(* IEC 61131-3 sources: plcassist-cli/packages/volt-lsp-iec/test-corpus/bakon-nano/Device/Plc Logic/Application/Library Manager/CmpBinTagUtilIec, 34 files *)

(* ---- BTAGALIGNMENTS.gvl ---- *)
VAR_GLOBAL
	ALIGN42 : BTagAlignment := STRUCT(uiModulus := 4, uiRemainder := 2);
	ALIGN40 : BTagAlignment := STRUCT(uiModulus := 4, uiRemainder := 0);
END_VAR

(* ---- RETURNVALUES.gvl ---- *)
VAR_GLOBAL
	ERR_OK : UDINT := 16#0;
	ERR_FAILED : UDINT := 16#1;
	ERR_PARAMETER : UDINT := 16#2;
	ERR_NOTIMPLEMENTED : UDINT := 16#C;
	ERR_NOMEMORY : UDINT := 16#11;
	ERR_BTAG_TAGOVERLAP : UDINT := 16#400;
	ERR_BTAG_BUFFEROVERRUN : UDINT := 16#401;
	ERR_BTAG_MAXNESTINGDEPTH : UDINT := 16#402;
	ERR_BTAG_NOTAG : UDINT := 16#403;
	ERR_BTAG_NODATATAG : UDINT := 16#404;
	ERR_BTAG_NOCONTAINERTAG : UDINT := 16#405;
	ERR_BTAG_NOTTOPLEVEL : UDINT := 16#406;
	ERR_BTAG_ALIGNMENT : UDINT := 16#407;
	INVALID_HANDLE : __UXINT := RTS_INVALID_HANDLE;
END_VAR

(* ---- BTAGREADERCREATE.fun ---- *)
FUNCTION BTAGREADERCREATE : RTS_IEC_HANDLE
VAR_INPUT
	PBUFFER : POINTER TO BYTE;
	DWSIZE : DWORD;
	PRESULT : POINTER TO RTS_IEC_RESULT;
END_VAR
END_FUNCTION

(* ---- BTAGREADERCREATEDYNAMIC.fun ---- *)
FUNCTION BTAGREADERCREATEDYNAMIC : RTS_IEC_HANDLE
VAR_INPUT
	PRESULT : POINTER TO RTS_IEC_RESULT;
END_VAR
END_FUNCTION

(* ---- BTAGREADERDESTROY.fun ---- *)
FUNCTION BTAGREADERDESTROY : RTS_IEC_RESULT
VAR_INPUT
	HREADER : RTS_IEC_HANDLE;
END_VAR
END_FUNCTION

(* ---- BTAGREADERGETCOMPLEXCONTENT.fun ---- *)
FUNCTION BTAGREADERGETCOMPLEXCONTENT : RTS_IEC_RESULT
VAR_INPUT
	HREADER : RTS_IEC_HANDLE;
	PPBUFFER : POINTER TO POINTER TO BYTE;
	PULSIZE : POINTER TO UDINT;
END_VAR
END_FUNCTION

(* ---- BTAGREADERGETCONTENT.fun ---- *)
FUNCTION BTAGREADERGETCONTENT : RTS_IEC_RESULT
VAR_INPUT
	HREADER : RTS_IEC_HANDLE;
	PPBUFFER : POINTER TO POINTER TO BYTE;
	PULSIZE : POINTER TO UDINT;
END_VAR
END_FUNCTION

(* ---- BTAGREADERGETSTRING.fun ---- *)
FUNCTION BTAGREADERGETSTRING : RTS_IEC_RESULT
VAR_INPUT
	HREADER : RTS_IEC_HANDLE;
	PPBUFFER : POINTER TO POINTER TO BYTE;
	PULSIZE : POINTER TO UDINT;
	BADDENDOFSTRING : BOOL;
END_VAR
END_FUNCTION

(* ---- BTAGREADERGETTAGID.fun ---- *)
FUNCTION BTAGREADERGETTAGID : RTS_IEC_RESULT
VAR_INPUT
	HREADER : RTS_IEC_HANDLE;
	PULTAGID : POINTER TO UDINT;
END_VAR
END_FUNCTION

(* ---- BTAGREADERGETTAGLEN.fun ---- *)
FUNCTION BTAGREADERGETTAGLEN : RTS_IEC_RESULT
VAR_INPUT
	HREADER : RTS_IEC_HANDLE;
	PULTAGLEN : POINTER TO UDINT;
END_VAR
END_FUNCTION

(* ---- BTAGREADERINIT.fun ---- *)
FUNCTION BTAGREADERINIT : RTS_IEC_RESULT
VAR_INPUT
	HREADER : RTS_IEC_HANDLE;
	PBUFFER : POINTER TO BYTE;
	DWBUFFERSIZE : DWORD;
END_VAR
END_FUNCTION

(* ---- BTAGREADERISDATATAG.fun ---- *)
FUNCTION BTAGREADERISDATATAG : RTS_IEC_RESULT
VAR_INPUT
	HREADER : RTS_IEC_HANDLE;
	PBDATATAG : POINTER TO BOOL;
END_VAR
END_FUNCTION

(* ---- BTAGREADERMOVENEXT.fun ---- *)
FUNCTION BTAGREADERMOVENEXT : RTS_IEC_RESULT
VAR_INPUT
	HREADER : RTS_IEC_HANDLE;
	PNELEMENTTYPE : POINTER TO BTagElementType;
END_VAR
END_FUNCTION

(* ---- BTAGREADERPEEKNEXT.fun ---- *)
FUNCTION BTAGREADERPEEKNEXT : BTagElementType
VAR_INPUT
	HREADER : RTS_IEC_HANDLE;
END_VAR
END_FUNCTION

(* ---- BTAGREADERSKIPCONTENT.fun ---- *)
FUNCTION BTAGREADERSKIPCONTENT : RTS_IEC_RESULT
VAR_INPUT
	HREADER : RTS_IEC_HANDLE;
END_VAR
END_FUNCTION

(* ---- BTAGSWAPHEADER.fun ---- *)
FUNCTION BTAGSWAPHEADER : DWORD
VAR_INPUT
	PHEADERTAG : POINTER TO DWORD;
	BSWAP : DINT;
END_VAR
END_FUNCTION

(* ---- BTAGWRITERAPPENDBLOB.fun ---- *)
FUNCTION BTAGWRITERAPPENDBLOB : RTS_IEC_RESULT
VAR_INPUT
	HWRITER : RTS_IEC_HANDLE;
	PDATA : POINTER TO BYTE;
	DWDATASIZE : DWORD;
END_VAR
END_FUNCTION

(* ---- BTAGWRITERAPPENDDUMMYBYTES.fun ---- *)
FUNCTION BTAGWRITERAPPENDDUMMYBYTES : RTS_IEC_RESULT
VAR_INPUT
	HWRITER : RTS_IEC_HANDLE;
	BTFILL : BYTE;
	ULCOUNT : DWORD;
END_VAR
END_FUNCTION

(* ---- BTAGWRITERAPPENDFILLBYTES.fun ---- *)
FUNCTION BTAGWRITERAPPENDFILLBYTES : RTS_IEC_RESULT
VAR_INPUT
	HWRITER : RTS_IEC_HANDLE;
	BTFILL : BYTE;
	ALIGNMENT : BTagAlignment;
END_VAR
END_FUNCTION

(* ---- BTAGWRITERAPPENDRAW.fun ---- *)
FUNCTION BTAGWRITERAPPENDRAW : RTS_IEC_RESULT
VAR_INPUT
	HWRITER : RTS_IEC_HANDLE;
	PPDATA : POINTER TO POINTER TO BYTE;
	DWSIZE : DWORD;
END_VAR
END_FUNCTION

(* ---- BTAGWRITERAPPENDWSTRING.fun ---- *)
FUNCTION BTAGWRITERAPPENDWSTRING : RTS_IEC_RESULT
VAR_INPUT
	HWRITER : RTS_IEC_HANDLE;
	WSZSTRING : REFERENCE TO WSTRING;
END_VAR
END_FUNCTION

(* ---- BTAGWRITERCREATE.fun ---- *)
FUNCTION BTAGWRITERCREATE : RTS_IEC_HANDLE
VAR_INPUT
	PBUFFER : POINTER TO BYTE;
	DWSIZE : DWORD;
	PRESULT : POINTER TO RTS_IEC_RESULT;
END_VAR
END_FUNCTION

(* ---- BTAGWRITERCREATEDYNAMIC.fun ---- *)
FUNCTION BTAGWRITERCREATEDYNAMIC : RTS_IEC_HANDLE
VAR_INPUT
	PRESULT : POINTER TO RTS_IEC_RESULT;
END_VAR
END_FUNCTION

(* ---- BTAGWRITERCREATESAVEPOINT.fun ---- *)
FUNCTION BTAGWRITERCREATESAVEPOINT : RTS_IEC_HANDLE
VAR_INPUT
	HWRITER : RTS_IEC_HANDLE;
	PDATA : POINTER TO BYTE;
	DWDATASIZE : DWORD;
	PRESULT : POINTER TO RTS_IEC_RESULT;
END_VAR
END_FUNCTION

(* ---- BTAGWRITERCREATESAVEPOINTDYNAMIC.fun ---- *)
FUNCTION BTAGWRITERCREATESAVEPOINTDYNAMIC : RTS_IEC_HANDLE
VAR_INPUT
	HWRITER : RTS_IEC_HANDLE;
	PRESULT : POINTER TO RTS_IEC_RESULT;
END_VAR
END_FUNCTION

(* ---- BTAGWRITERDESTROY.fun ---- *)
FUNCTION BTAGWRITERDESTROY : RTS_IEC_RESULT
VAR_INPUT
	HWRITER : RTS_IEC_HANDLE;
END_VAR
END_FUNCTION

(* ---- BTAGWRITERDESTROYSAVEPOINT.fun ---- *)
FUNCTION BTAGWRITERDESTROYSAVEPOINT : RTS_IEC_RESULT
VAR_INPUT
	HSAVEPOINT : RTS_IEC_HANDLE;
END_VAR
END_FUNCTION

(* ---- BTAGWRITERENDTAG.fun ---- *)
FUNCTION BTAGWRITERENDTAG : RTS_IEC_RESULT
VAR_INPUT
	HWRITER : RTS_IEC_HANDLE;
	UDITAGID : UDINT;
END_VAR
END_FUNCTION

(* ---- BTAGWRITERFINISH.fun ---- *)
FUNCTION BTAGWRITERFINISH : RTS_IEC_RESULT
VAR_INPUT
	HWRITER : RTS_IEC_HANDLE;
	PPBUFFER : POINTER TO POINTER TO BYTE;
	PUISIZE : POINTER TO UDINT;
END_VAR
END_FUNCTION

(* ---- BTAGWRITERINIT.fun ---- *)
FUNCTION BTAGWRITERINIT : RTS_IEC_RESULT
VAR_INPUT
	HWRITER : RTS_IEC_HANDLE;
	PBUFFER : POINTER TO BYTE;
	DWBUFFERSIZE : DWORD;
END_VAR
END_FUNCTION

(* ---- BTAGWRITERINIT2.fun ---- *)
FUNCTION BTAGWRITERINIT2 : RTS_IEC_RESULT
VAR_INPUT
	HWRITER : RTS_IEC_HANDLE;
	PBUFFER : POINTER TO BYTE;
	DWBUFFERSIZE : DWORD;
	BSWAP : DINT;
END_VAR
END_FUNCTION

(* ---- BTAGWRITERRESTORESAVEPOINT.fun ---- *)
FUNCTION BTAGWRITERRESTORESAVEPOINT : RTS_IEC_RESULT
VAR_INPUT
	HWRITER : RTS_IEC_HANDLE;
	HSAVEPOINT : RTS_IEC_HANDLE;
END_VAR
END_FUNCTION

(* ---- BTAGWRITERSTARTTAG.fun ---- *)
FUNCTION BTAGWRITERSTARTTAG : RTS_IEC_RESULT
VAR_INPUT
	HWRITER : RTS_IEC_HANDLE;
	UDITAGID : UDINT;
	ALIGNMENT : BTagAlignment;
	UDIMINLENGTHSIZE : UDINT;
END_VAR
END_FUNCTION

(* ---- BTAGWRITERSWITCHBUFFER.fun ---- *)
FUNCTION BTAGWRITERSWITCHBUFFER : RTS_IEC_RESULT
VAR_INPUT
	HWRITER : RTS_IEC_HANDLE;
	PNEWBUFFER : POINTER TO BYTE;
	DWNEWBUFFERSIZE : DWORD;
	PPOLDBUFFER : POINTER TO POINTER TO BYTE;
END_VAR
END_FUNCTION
